Universal Robots URScript: T001_codellama_34b_adversarial_A8.5_rep1.urscript

def simple_pick_place(payload):
    # Move to home position
    movej(p[0, 0, 0, 0, 0, 0], v=200.0)

    # Approach pick point
    movel(p[0, 0, -150, 0, 0, 0], v=200.0)

    # Descend
